(* IEC 61131-3 sources: stf-hw/web/public/sil (part 3) *)

CONFIGURATION Cell
    RESOURCE Plc ON PLC
        TASK Scan(INTERVAL := T#5MS, PRIORITY := 0);
        PROGRAM Run WITH Scan : MAIN;
    END_RESOURCE
END_CONFIGURATION
